DATA_BLOCK "GDB_FraktalMain"
{ S7_Optimized_Access := 'TRUE' }
VERSION : 0.1
NON_RETAIN
"FB_FraktalMain"
BEGIN
END_DATA_BLOCK
